TYPE ST_TwoHandControl :
STRUCT
	diButton1		 AT %I* : BOOL;
	diStartButton	 AT %I* : BOOL;
	diStopButton	 AT %I* : BOOL;
	diTwoHand		 AT %I* : BOOL;
	diTwoHand1		 AT %I* : BOOL;
	diTwoHand2		 AT %I* : BOOL;
	diSafetySwitch	 AT %I* : BOOL;
	doStartLED		 AT %Q* : BOOL;
	doStopLED		 AT %Q* : BOOL;
	
	xButton1RTrigger		: BOOL;
	xButton1FTrigger		: BOOL;
	xStartRTrigger			: BOOL;
	xStartFTrigger			: BOOL;
	xStopRTrigger			: BOOL;
	xStopFTrigger			: BOOL;
	xTwoHandRTrigger		: BOOL;
	xTwoHandFTRigger		: BOOL;
	xSafetySwitchRTrigger	: BOOL;
	xSafetySwitchFTrigger	: BOOL;
	xStopButtonDelayTrigger	: BOOL;
END_STRUCT
END_TYPE

(* stored: Version 1.1.0.1, ProductVersion 3.1.4024.12
   DUT ST_TwoHandControl: Id {819477b7-5f09-4f80-b3d0-b8b206edd0cb} *)
